Fanuc KAREL source: KD00037.KL

PROGRAM KD00037
%NOLOCKGROUP
VAR
  I: INTEGER
  J: INTEGER
  B: BOOLEAN
  R: REAL
  S: STRING[80]
BEGIN
  CONDITION[1]:
  WHEN DIN[1] = ON DO
    UNPAUSE
  ENDCONDITION
END KD00037
